SUBAPPLICATION Sperrblock_Button_OR8_TO_logiBUS_QXA_BG (* Sperrblock: Button ODER 8 Anforderungen auf logiBUS-Ausgang, Hintergrundfarbe Gruen/Weiss *)
  (* Standard: 61499-2; Description: Copyright (c) 2026 Meisterschulen am Ostbahnhof This program and the accompanying materials are made available under the terms of the Eclipse Public License 2.0 which is available at https://www.eclipse.org/legal/epl-2.0/ SPDX-License-Identifier: EPL-2.0 *)
  (* Version 1.0, 2026-10-31, Franz Höpfinger, Meisterschulen am Ostbahnhof, Aus Getreidehacke func/Manual/SB in MyLib::sys verschoben und umbenannt, INIT/INITO/QI/QO ergaenzt, Output als Parameter (vorher fest Output_Q2). *)
  PACKAGE MyLib::sys;
  IMPORT isobus::UT::Q::const::IDs::ID_NULL;
  IMPORT logiBUS::io::DQ::logiBUS_DO;
  IMPORT logiBUS::io::DQ::logiBUS_DO_S;
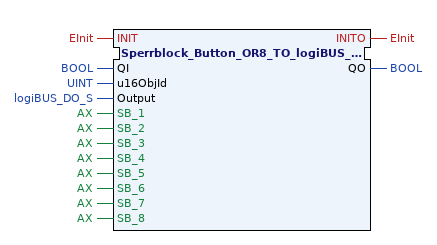
  EVENT_INPUT
    INIT : EInit; (* Initialization Request *)
  END_EVENT
  EVENT_OUTPUT
    INITO : EInit; (* Initialization Confirm *)
  END_EVENT
  VAR_INPUT
    QI : BOOL := TRUE; (* Quality Input - TRUE to enable service *)
    u16ObjId : UINT := ID_NULL; (* Object ID Button Sperrblock *)
    Output : logiBUS::io::DQ::logiBUS_DO_S := logiBUS_DO::Invalid; (* logiBUS-Ausgang Sperrblock *)
  END_VAR
  VAR_OUTPUT
    QO : BOOL; (* Quality Output - TRUE if service executed successfully *)
  END_VAR
  SOCKETS
    SB_1 : adapter::types::unidirectional::AX; (* Anforderung Sperrblock 1 *)
    SB_2 : adapter::types::unidirectional::AX; (* Anforderung Sperrblock 2 *)
    SB_3 : adapter::types::unidirectional::AX; (* Anforderung Sperrblock 3 *)
    SB_4 : adapter::types::unidirectional::AX; (* Anforderung Sperrblock 4 *)
    SB_5 : adapter::types::unidirectional::AX; (* Anforderung Sperrblock 5 *)
    SB_6 : adapter::types::unidirectional::AX; (* Anforderung Sperrblock 6 *)
    SB_7 : adapter::types::unidirectional::AX; (* Anforderung Sperrblock 7 *)
    SB_8 : adapter::types::unidirectional::AX; (* Anforderung Sperrblock 8 *)
  END_SOCKETS
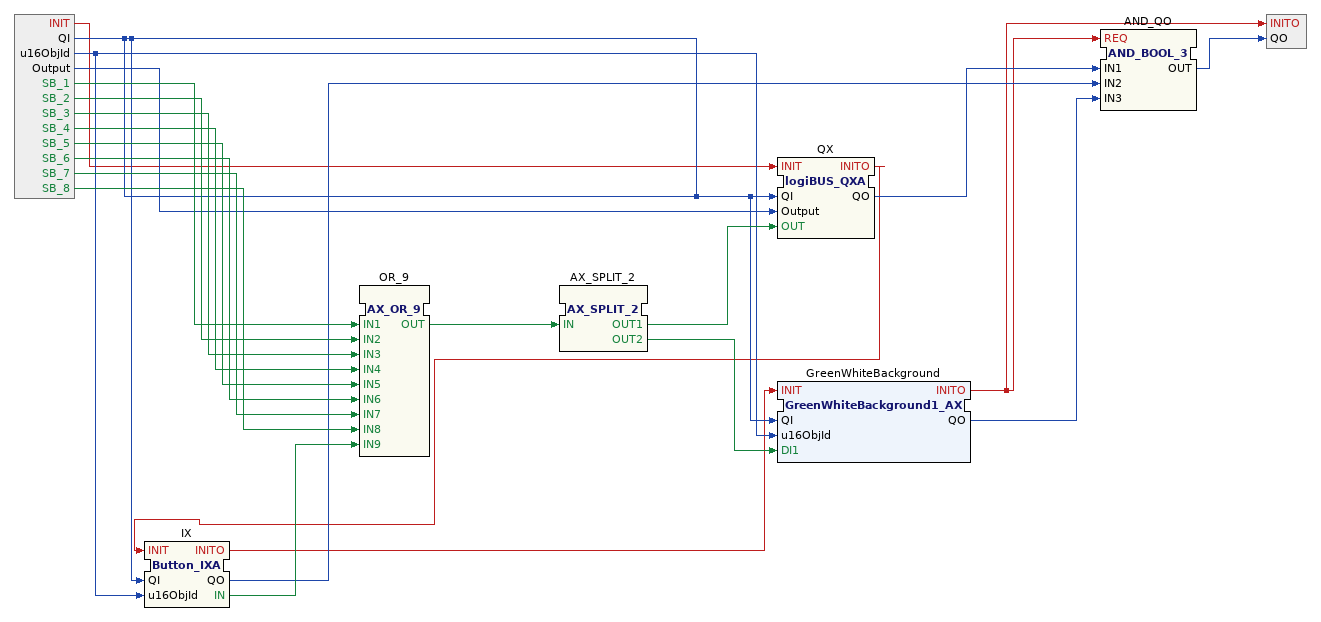
  FBS
    IX : isobus::UT::io::Button::Button_IXA;
    OR_9 : adapter::booleanOperators::AX_OR_9;
    AX_SPLIT_2 : adapter::events::unidirectional::AX_SPLIT_2;
    QX : logiBUS::io::DQ::logiBUS_QXA;
    AND_QO : iec61131::booleanOperators::AND_BOOL_3;
  END_FBS
  SUBAPPS
    GreenWhiteBackground : MyLib::sys::GreenWhiteBackground1_AX;
  END_SUBAPPS
  EVENT_CONNECTIONS
    INIT TO QX.INIT;
    QX.INITO TO IX.INIT;
    IX.INITO TO GreenWhiteBackground.INIT;
    GreenWhiteBackground.INITO TO INITO;
    GreenWhiteBackground.INITO TO AND_QO.REQ;
  END_CONNECTIONS
  DATA_CONNECTIONS
    QI TO QX.QI;
    QI TO IX.QI;
    QI TO GreenWhiteBackground.QI;
    u16ObjId TO IX.u16ObjId;
    u16ObjId TO GreenWhiteBackground.u16ObjId;
    Output TO QX.Output;
    QX.QO TO AND_QO.IN1;
    IX.QO TO AND_QO.IN2;
    GreenWhiteBackground.QO TO AND_QO.IN3;
    AND_QO.OUT TO QO;
  END_CONNECTIONS
  ADAPTER_CONNECTIONS
    SB_1 TO OR_9.IN1;
    SB_2 TO OR_9.IN2;
    SB_3 TO OR_9.IN3;
    SB_4 TO OR_9.IN4;
    SB_5 TO OR_9.IN5;
    SB_6 TO OR_9.IN6;
    SB_7 TO OR_9.IN7;
    SB_8 TO OR_9.IN8;
    IX.IN TO OR_9.IN9;
    OR_9.OUT TO AX_SPLIT_2.IN;
    AX_SPLIT_2.OUT1 TO QX.OUT;
    AX_SPLIT_2.OUT2 TO GreenWhiteBackground.DI1;
  END_CONNECTIONS
END_SUBAPPLICATION
